Fanuc KAREL source: KT00855.KL

PROGRAM KT00855
%NOLOCKGROUP
VAR
  S1: STRING[80]
  S2: STRING[80]
  OUT: REAL
BEGIN
  S1 = 'A'
  S2 = 'B'
  S1 = 'A'
  S2 = 'B'
  OUT = TAN(S1)
END KT00855
